TYPE "DT_REGULATOR_INTERFACE_ALL"
VERSION : 0.1
   STRUCT
      WATER_LEVEL : "DT_REGULATOR_INTERFACE";
      GATE_1 : "DT_REGULATOR_INTERFACE";
      GATE_2 : "DT_REGULATOR_INTERFACE";
      GATE_3 : "DT_REGULATOR_INTERFACE";
      GATE_4 : "DT_REGULATOR_INTERFACE";
      GATE_5 : "DT_REGULATOR_INTERFACE";
      GATE_6 : "DT_REGULATOR_INTERFACE";
      GATE_7 : "DT_REGULATOR_INTERFACE";
      GATE_8 : "DT_REGULATOR_INTERFACE";
      GATE_9 : "DT_REGULATOR_INTERFACE";
      GATE_10 : "DT_REGULATOR_INTERFACE";
      SPARE_11 : "DT_REGULATOR_INTERFACE";
      SPARE_12 : "DT_REGULATOR_INTERFACE";
      SPARE_13 : "DT_REGULATOR_INTERFACE";
      SPARE_14 : "DT_REGULATOR_INTERFACE";
      SPARE_15 : "DT_REGULATOR_INTERFACE";
      SPARE_16 : "DT_REGULATOR_INTERFACE";
      SPARE_17 : "DT_REGULATOR_INTERFACE";
      SPARE_18 : "DT_REGULATOR_INTERFACE";
      SPARE_19 : "DT_REGULATOR_INTERFACE";
      SPARE_20 : "DT_REGULATOR_INTERFACE";
      SPARE_21 : "DT_REGULATOR_INTERFACE";
      SPARE_22 : "DT_REGULATOR_INTERFACE";
      SPARE_23 : "DT_REGULATOR_INTERFACE";
      SPARE_24 : "DT_REGULATOR_INTERFACE";
      SPARE_25 : "DT_REGULATOR_INTERFACE";
      SPARE_26 : "DT_REGULATOR_INTERFACE";
      SPARE_27 : "DT_REGULATOR_INTERFACE";
      SPARE_28 : "DT_REGULATOR_INTERFACE";
      SPARE_29 : "DT_REGULATOR_INTERFACE";
      SPARE_30 : "DT_REGULATOR_INTERFACE";
      SPARE_31 : "DT_REGULATOR_INTERFACE";
   END_STRUCT;

END_TYPE

